FUNCTION_BLOCK ButtonPanel_Control (* Extracted Composite Function Block Type *)
  (* Standard: 61499-2 *)
  (* Version 10/19/2026, lizar *)
  PACKAGE Main;
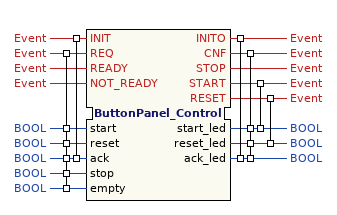
  EVENT_INPUT
    INIT WITH ack; (* Event input *)
    REQ WITH start, reset, stop, ack, empty; (* Normal Execution Request *)
    READY;
    NOT_READY;
  END_EVENT
  EVENT_OUTPUT
    INITO WITH ack_led;
    CNF WITH start_led, reset_led, ack_led; (* Execution Confirmation *)
    STOP;
    START WITH start_led;
    RESET WITH reset_led;
  END_EVENT
  VAR_INPUT
    start : BOOL;
    reset : BOOL;
    ack : BOOL; (* Event permission *)
    stop : BOOL;
    empty : BOOL;
  END_VAR
  VAR_OUTPUT
    start_led : BOOL;
    reset_led : BOOL;
    ack_led : BOOL; (* Output event qualifier *)
  END_VAR
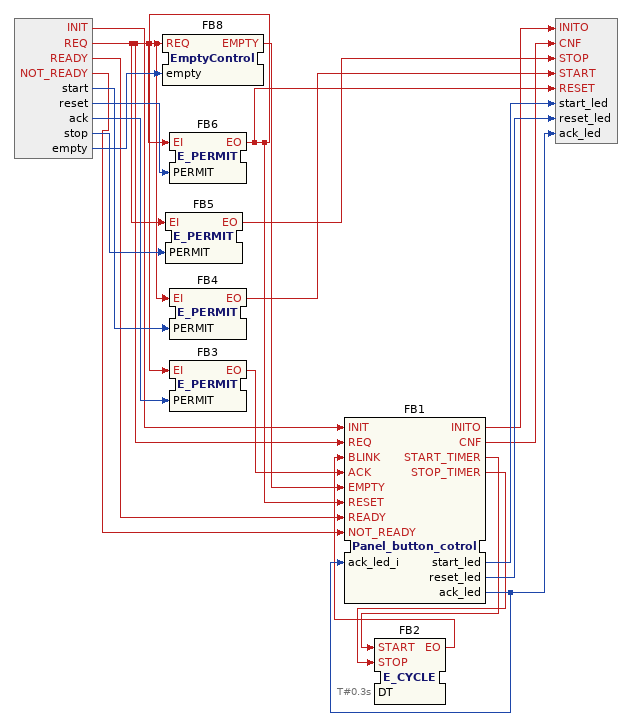
  FBS
    FB1 : Panel_button_cotrol;
    FB2 : E_CYCLE(DT := T#0.3s);
    FB3 : E_PERMIT;
    FB4 : E_PERMIT;
    FB5 : E_PERMIT;
    FB6 : E_PERMIT;
    FB8 : EmptyControl;
  END_FBS
  EVENT_CONNECTIONS
    FB1.START_TIMER TO FB2.START;
    FB1.STOP_TIMER TO FB2.STOP;
    FB2.EO TO FB1.BLINK;
    FB3.EO TO FB1.ACK;
    REQ TO FB1.REQ;
    FB1.CNF TO CNF;
    REQ TO FB3.EI;
    REQ TO FB4.EI;
    FB4.EO TO START;
    INIT TO FB1.INIT;
    FB1.INITO TO INITO;
    REQ TO FB5.EI;
    FB5.EO TO STOP;
    FB6.EO TO RESET;
    REQ TO FB6.EI;
    FB6.EO TO FB1.RESET;
    READY TO FB1.READY;
    NOT_READY TO FB1.NOT_READY;
    FB6.EO TO FB8.REQ;
    FB8.EMPTY TO FB1.EMPTY;
    REQ TO FB8.REQ;
  END_CONNECTIONS
  DATA_CONNECTIONS
    ack TO FB3.PERMIT;
    FB1.start_led TO start_led;
    FB1.reset_led TO reset_led;
    FB1.ack_led TO ack_led;
    FB1.ack_led TO FB1.ack_led_i;
    start TO FB4.PERMIT;
    stop TO FB5.PERMIT;
    reset TO FB6.PERMIT;
    empty TO FB8.empty;
  END_CONNECTIONS
END_FUNCTION_BLOCK
